(* IEC 61131-3 sources: rusty/tests/lit/cfc/variables/literal_assignment, 1 file *)

(* ---- main.st ---- *)
FUNCTION main : DINT
    literal_assignment();
    // CHECK: x = 42
    printf('x = %d$N', literal_assignment.x);
END_FUNCTION
